{attribute 'Tc2GvlVarNames'}
VAR_GLOBAL CONSTANT
	usnFileArrayMaxDimR					:USINT := 100;		(* 0..usnMaxDimR - Number of rows to read. *)
	usnFileArrayMaxDimC					:USINT := 4;  		(* 0..usnMaxDimC -  Number of columns to read. *)
END_VAR

(* stored: Version 1.1.0.1, ProductVersion 3.1.4024.15
   GVL GVL_FB_LoadFromFile_1: Id {050184dd-a766-4925-a427-e29cf8bda48a} *)
